// TIA Portal V20 export
Screen "Pop-up_ALARM_HISTORY_LEGEND_Popup"  330x100
  ScreenItem "Background" at 0,0 size 330x100  Type=HmiRectangle
  ScreenItem "Textfeld_Legende" at 1,1 size 328x25  Type=HmiTextBox
  ScreenItem "Textfeld_11" at 10,33 size 230x60  Type=HmiTextBox
  ScreenItem "Cancel Mode" at 239,1 size 90x60  Type=HmiButton
